// TIA Portal V21 export
DATA_BLOCK "IDB_AnaTimerCaller"   // DB15
// stored: InstanceOfName FB_AnaTimerCaller, InstanceOfType FB
"FB_AnaTimerCaller"
   // VAR_INPUT
   //    Enable : Bool;
   //    Start : Bool;
   // END_VAR
   // VAR_OUTPUT
   //    Done : Bool;
   // END_VAR
   // VAR
   //    Inner { S7_SetPoint := 'True'} : "FB_AnaTimerInner";
   // END_VAR
BEGIN
END_DATA_BLOCK
